(* IEC 61131-3 sources: TIA2AX/tests/V18/test_projects/expected/HW_Plc1518V3_CmmtAs/PLC_LINE, 7 files *)

(* ---- HwIdentifiers.st ---- *)
TYPE
	HwIdentifiers : WORD
	(
		PLC_LINE_Rail_0 :=	WORD#256,
		PLC_LINE :=	WORD#48,
		PLC_LINE_Card_reader_writer_1 :=	WORD#51,
		PLC_LINE_CPU_display_1 :=	WORD#54,
		PLC_LINE_OPC_UA_1 :=	WORD#117,
		PLC_LINE_PROFINET_interface_1 :=	WORD#64,
		PLC_LINE_PROFINET_interface_1_Port_1 :=	WORD#65,
		PLC_LINE_PROFINET_interface_1_Port_2 :=	WORD#66,
		PLC_LINE_PROFINET_interface_2 :=	WORD#72,
		PLC_LINE_PROFINET_interface_2_Port_1 :=	WORD#73,
		PLC_LINE_DP_interface_1 :=	WORD#60,
		PLC_LINE_PROFINET_interface_GBIT_3 :=	WORD#120,
		PLC_LINE_PROFINET_interface_GBIT_3_Port_1 :=	WORD#121,
		cmmtas_PN_IO_Interface :=	WORD#271,
		cmmtas_PN_IO_Interface_Port_1 :=	WORD#260,
		cmmtas_PN_IO_Interface_Port_2 :=	WORD#261,
		cmmtas_CMMT_AS_MP :=	WORD#272,
		cmmtas_DO_SERVO_1_Module_Access_Point :=	WORD#264,
		cmmtas_DO_SERVO_1_Siemens_telegram_111_PZD_12_12 :=	WORD#265,
		cmmtas_DO_SERVO_1_Siemens_telegram_750_PZD_4_1 :=	WORD#266,
		cmmtas_Siemens_telegram_111_PZD_12_12 :=	WORD#265,
		cmmtas_Siemens_telegram_750_PZD_4_1 :=	WORD#266,
		NONE:= WORD#0
	);
END_TYPE

(* ---- HwInputs.st ---- *)
TYPE
	HwInputs : STRUCT
		cmmtas_DO_SERVO_1_Siemens_telegram_111_PZD_12_12 AT %B100 : ARRAY[0..23] OF BYTE;
		cmmtas_DO_SERVO_1_Siemens_telegram_750_PZD_4_1 AT %B124 : WORD;
	END_STRUCT;
END_TYPE

(* ---- HwOutputs.st ---- *)
TYPE
	HwOutputs : STRUCT
		cmmtas_DO_SERVO_1_Siemens_telegram_111_PZD_12_12 AT %B100 : ARRAY[0..23] OF BYTE;
		cmmtas_DO_SERVO_1_Siemens_telegram_750_PZD_4_1 AT %B124 : ARRAY[0..7] OF BYTE;
	END_STRUCT;
END_TYPE

(* ---- PlcInputs.st ---- *)
TYPE
	PlcInputs : STRUCT
		cmmtas_DO_SERVO_1_Siemens_telegram_111_PZD_12_12 : ARRAY[0..23] OF BYTE;
		cmmtas_DO_SERVO_1_Siemens_telegram_750_PZD_4_1 : WORD;
	END_STRUCT;
END_TYPE

(* ---- PlcOutputs.st ---- *)
TYPE
	PlcOutputs : STRUCT
		cmmtas_DO_SERVO_1_Siemens_telegram_111_PZD_12_12 : ARRAY[0..23] OF BYTE;
		cmmtas_DO_SERVO_1_Siemens_telegram_750_PZD_4_1 : ARRAY[0..7] OF BYTE;
	END_STRUCT;
END_TYPE

(* ---- CopyInputs.st ---- *)
FUNCTION CopyInputs
	VAR_EXTERNAL
		HwInputs : HwInputs;
		PlcInputs : PlcInputs;
	END_VAR
	PlcInputs.cmmtas_DO_SERVO_1_Siemens_telegram_111_PZD_12_12[0] := HwInputs.cmmtas_DO_SERVO_1_Siemens_telegram_111_PZD_12_12[0];
	PlcInputs.cmmtas_DO_SERVO_1_Siemens_telegram_111_PZD_12_12[1] := HwInputs.cmmtas_DO_SERVO_1_Siemens_telegram_111_PZD_12_12[1];
	PlcInputs.cmmtas_DO_SERVO_1_Siemens_telegram_111_PZD_12_12[2] := HwInputs.cmmtas_DO_SERVO_1_Siemens_telegram_111_PZD_12_12[2];
	PlcInputs.cmmtas_DO_SERVO_1_Siemens_telegram_111_PZD_12_12[3] := HwInputs.cmmtas_DO_SERVO_1_Siemens_telegram_111_PZD_12_12[3];
	PlcInputs.cmmtas_DO_SERVO_1_Siemens_telegram_111_PZD_12_12[4] := HwInputs.cmmtas_DO_SERVO_1_Siemens_telegram_111_PZD_12_12[4];
	PlcInputs.cmmtas_DO_SERVO_1_Siemens_telegram_111_PZD_12_12[5] := HwInputs.cmmtas_DO_SERVO_1_Siemens_telegram_111_PZD_12_12[5];
	PlcInputs.cmmtas_DO_SERVO_1_Siemens_telegram_111_PZD_12_12[6] := HwInputs.cmmtas_DO_SERVO_1_Siemens_telegram_111_PZD_12_12[6];
	PlcInputs.cmmtas_DO_SERVO_1_Siemens_telegram_111_PZD_12_12[7] := HwInputs.cmmtas_DO_SERVO_1_Siemens_telegram_111_PZD_12_12[7];
	PlcInputs.cmmtas_DO_SERVO_1_Siemens_telegram_111_PZD_12_12[8] := HwInputs.cmmtas_DO_SERVO_1_Siemens_telegram_111_PZD_12_12[8];
	PlcInputs.cmmtas_DO_SERVO_1_Siemens_telegram_111_PZD_12_12[9] := HwInputs.cmmtas_DO_SERVO_1_Siemens_telegram_111_PZD_12_12[9];
	PlcInputs.cmmtas_DO_SERVO_1_Siemens_telegram_111_PZD_12_12[10] := HwInputs.cmmtas_DO_SERVO_1_Siemens_telegram_111_PZD_12_12[10];
	PlcInputs.cmmtas_DO_SERVO_1_Siemens_telegram_111_PZD_12_12[11] := HwInputs.cmmtas_DO_SERVO_1_Siemens_telegram_111_PZD_12_12[11];
	PlcInputs.cmmtas_DO_SERVO_1_Siemens_telegram_111_PZD_12_12[12] := HwInputs.cmmtas_DO_SERVO_1_Siemens_telegram_111_PZD_12_12[12];
	PlcInputs.cmmtas_DO_SERVO_1_Siemens_telegram_111_PZD_12_12[13] := HwInputs.cmmtas_DO_SERVO_1_Siemens_telegram_111_PZD_12_12[13];
	PlcInputs.cmmtas_DO_SERVO_1_Siemens_telegram_111_PZD_12_12[14] := HwInputs.cmmtas_DO_SERVO_1_Siemens_telegram_111_PZD_12_12[14];
	PlcInputs.cmmtas_DO_SERVO_1_Siemens_telegram_111_PZD_12_12[15] := HwInputs.cmmtas_DO_SERVO_1_Siemens_telegram_111_PZD_12_12[15];
	PlcInputs.cmmtas_DO_SERVO_1_Siemens_telegram_111_PZD_12_12[16] := HwInputs.cmmtas_DO_SERVO_1_Siemens_telegram_111_PZD_12_12[16];
	PlcInputs.cmmtas_DO_SERVO_1_Siemens_telegram_111_PZD_12_12[17] := HwInputs.cmmtas_DO_SERVO_1_Siemens_telegram_111_PZD_12_12[17];
	PlcInputs.cmmtas_DO_SERVO_1_Siemens_telegram_111_PZD_12_12[18] := HwInputs.cmmtas_DO_SERVO_1_Siemens_telegram_111_PZD_12_12[18];
	PlcInputs.cmmtas_DO_SERVO_1_Siemens_telegram_111_PZD_12_12[19] := HwInputs.cmmtas_DO_SERVO_1_Siemens_telegram_111_PZD_12_12[19];
	PlcInputs.cmmtas_DO_SERVO_1_Siemens_telegram_111_PZD_12_12[20] := HwInputs.cmmtas_DO_SERVO_1_Siemens_telegram_111_PZD_12_12[20];
	PlcInputs.cmmtas_DO_SERVO_1_Siemens_telegram_111_PZD_12_12[21] := HwInputs.cmmtas_DO_SERVO_1_Siemens_telegram_111_PZD_12_12[21];
	PlcInputs.cmmtas_DO_SERVO_1_Siemens_telegram_111_PZD_12_12[22] := HwInputs.cmmtas_DO_SERVO_1_Siemens_telegram_111_PZD_12_12[22];
	PlcInputs.cmmtas_DO_SERVO_1_Siemens_telegram_111_PZD_12_12[23] := HwInputs.cmmtas_DO_SERVO_1_Siemens_telegram_111_PZD_12_12[23];
	PlcInputs.cmmtas_DO_SERVO_1_Siemens_telegram_750_PZD_4_1 := HwInputs.cmmtas_DO_SERVO_1_Siemens_telegram_750_PZD_4_1;
END_FUNCTION

(* ---- CopyOutputs.st ---- *)
FUNCTION CopyOutputs
	VAR_EXTERNAL
		HwOutputs : HwOutputs;
		PlcOutputs : PlcOutputs;
	END_VAR
	HwOutputs.cmmtas_DO_SERVO_1_Siemens_telegram_111_PZD_12_12[0] := PlcOutputs.cmmtas_DO_SERVO_1_Siemens_telegram_111_PZD_12_12[0];
	HwOutputs.cmmtas_DO_SERVO_1_Siemens_telegram_111_PZD_12_12[1] := PlcOutputs.cmmtas_DO_SERVO_1_Siemens_telegram_111_PZD_12_12[1];
	HwOutputs.cmmtas_DO_SERVO_1_Siemens_telegram_111_PZD_12_12[2] := PlcOutputs.cmmtas_DO_SERVO_1_Siemens_telegram_111_PZD_12_12[2];
	HwOutputs.cmmtas_DO_SERVO_1_Siemens_telegram_111_PZD_12_12[3] := PlcOutputs.cmmtas_DO_SERVO_1_Siemens_telegram_111_PZD_12_12[3];
	HwOutputs.cmmtas_DO_SERVO_1_Siemens_telegram_111_PZD_12_12[4] := PlcOutputs.cmmtas_DO_SERVO_1_Siemens_telegram_111_PZD_12_12[4];
	HwOutputs.cmmtas_DO_SERVO_1_Siemens_telegram_111_PZD_12_12[5] := PlcOutputs.cmmtas_DO_SERVO_1_Siemens_telegram_111_PZD_12_12[5];
	HwOutputs.cmmtas_DO_SERVO_1_Siemens_telegram_111_PZD_12_12[6] := PlcOutputs.cmmtas_DO_SERVO_1_Siemens_telegram_111_PZD_12_12[6];
	HwOutputs.cmmtas_DO_SERVO_1_Siemens_telegram_111_PZD_12_12[7] := PlcOutputs.cmmtas_DO_SERVO_1_Siemens_telegram_111_PZD_12_12[7];
	HwOutputs.cmmtas_DO_SERVO_1_Siemens_telegram_111_PZD_12_12[8] := PlcOutputs.cmmtas_DO_SERVO_1_Siemens_telegram_111_PZD_12_12[8];
	HwOutputs.cmmtas_DO_SERVO_1_Siemens_telegram_111_PZD_12_12[9] := PlcOutputs.cmmtas_DO_SERVO_1_Siemens_telegram_111_PZD_12_12[9];
	HwOutputs.cmmtas_DO_SERVO_1_Siemens_telegram_111_PZD_12_12[10] := PlcOutputs.cmmtas_DO_SERVO_1_Siemens_telegram_111_PZD_12_12[10];
	HwOutputs.cmmtas_DO_SERVO_1_Siemens_telegram_111_PZD_12_12[11] := PlcOutputs.cmmtas_DO_SERVO_1_Siemens_telegram_111_PZD_12_12[11];
	HwOutputs.cmmtas_DO_SERVO_1_Siemens_telegram_111_PZD_12_12[12] := PlcOutputs.cmmtas_DO_SERVO_1_Siemens_telegram_111_PZD_12_12[12];
	HwOutputs.cmmtas_DO_SERVO_1_Siemens_telegram_111_PZD_12_12[13] := PlcOutputs.cmmtas_DO_SERVO_1_Siemens_telegram_111_PZD_12_12[13];
	HwOutputs.cmmtas_DO_SERVO_1_Siemens_telegram_111_PZD_12_12[14] := PlcOutputs.cmmtas_DO_SERVO_1_Siemens_telegram_111_PZD_12_12[14];
	HwOutputs.cmmtas_DO_SERVO_1_Siemens_telegram_111_PZD_12_12[15] := PlcOutputs.cmmtas_DO_SERVO_1_Siemens_telegram_111_PZD_12_12[15];
	HwOutputs.cmmtas_DO_SERVO_1_Siemens_telegram_111_PZD_12_12[16] := PlcOutputs.cmmtas_DO_SERVO_1_Siemens_telegram_111_PZD_12_12[16];
	HwOutputs.cmmtas_DO_SERVO_1_Siemens_telegram_111_PZD_12_12[17] := PlcOutputs.cmmtas_DO_SERVO_1_Siemens_telegram_111_PZD_12_12[17];
	HwOutputs.cmmtas_DO_SERVO_1_Siemens_telegram_111_PZD_12_12[18] := PlcOutputs.cmmtas_DO_SERVO_1_Siemens_telegram_111_PZD_12_12[18];
	HwOutputs.cmmtas_DO_SERVO_1_Siemens_telegram_111_PZD_12_12[19] := PlcOutputs.cmmtas_DO_SERVO_1_Siemens_telegram_111_PZD_12_12[19];
	HwOutputs.cmmtas_DO_SERVO_1_Siemens_telegram_111_PZD_12_12[20] := PlcOutputs.cmmtas_DO_SERVO_1_Siemens_telegram_111_PZD_12_12[20];
	HwOutputs.cmmtas_DO_SERVO_1_Siemens_telegram_111_PZD_12_12[21] := PlcOutputs.cmmtas_DO_SERVO_1_Siemens_telegram_111_PZD_12_12[21];
	HwOutputs.cmmtas_DO_SERVO_1_Siemens_telegram_111_PZD_12_12[22] := PlcOutputs.cmmtas_DO_SERVO_1_Siemens_telegram_111_PZD_12_12[22];
	HwOutputs.cmmtas_DO_SERVO_1_Siemens_telegram_111_PZD_12_12[23] := PlcOutputs.cmmtas_DO_SERVO_1_Siemens_telegram_111_PZD_12_12[23];
	HwOutputs.cmmtas_DO_SERVO_1_Siemens_telegram_750_PZD_4_1[0] := PlcOutputs.cmmtas_DO_SERVO_1_Siemens_telegram_750_PZD_4_1[0];
	HwOutputs.cmmtas_DO_SERVO_1_Siemens_telegram_750_PZD_4_1[1] := PlcOutputs.cmmtas_DO_SERVO_1_Siemens_telegram_750_PZD_4_1[1];
	HwOutputs.cmmtas_DO_SERVO_1_Siemens_telegram_750_PZD_4_1[2] := PlcOutputs.cmmtas_DO_SERVO_1_Siemens_telegram_750_PZD_4_1[2];
	HwOutputs.cmmtas_DO_SERVO_1_Siemens_telegram_750_PZD_4_1[3] := PlcOutputs.cmmtas_DO_SERVO_1_Siemens_telegram_750_PZD_4_1[3];
	HwOutputs.cmmtas_DO_SERVO_1_Siemens_telegram_750_PZD_4_1[4] := PlcOutputs.cmmtas_DO_SERVO_1_Siemens_telegram_750_PZD_4_1[4];
	HwOutputs.cmmtas_DO_SERVO_1_Siemens_telegram_750_PZD_4_1[5] := PlcOutputs.cmmtas_DO_SERVO_1_Siemens_telegram_750_PZD_4_1[5];
	HwOutputs.cmmtas_DO_SERVO_1_Siemens_telegram_750_PZD_4_1[6] := PlcOutputs.cmmtas_DO_SERVO_1_Siemens_telegram_750_PZD_4_1[6];
	HwOutputs.cmmtas_DO_SERVO_1_Siemens_telegram_750_PZD_4_1[7] := PlcOutputs.cmmtas_DO_SERVO_1_Siemens_telegram_750_PZD_4_1[7];
END_FUNCTION
